RoboDK station: Robotic_Paint_Station.rdk

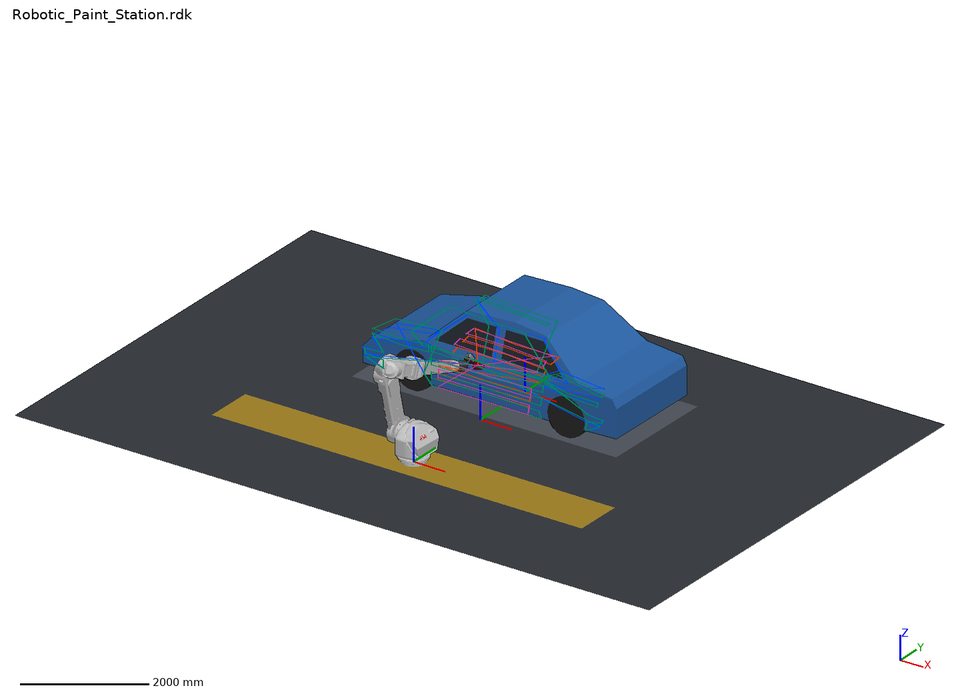
[picture v0: the station drawn from its stored meshes, robots at their saved joint values, targets as dots, program paths as lines]
Station Robotic_Paint_Station (saved by RoboDK 6.1.1). Poses are relative to the parent item; angles as X-Y-Z fixed-axis rotations.
  - frame ABB IRB 5500-27 Base at (0, 0, 0) mm
    - robot ABB IRB 5500-27: 6 axes, payload 16 kg, reach 2200 mm, repeatability 0.15 mm, weight 600 kg
        modified DH rows (alpha deg, a mm, theta deg, d mm): 0, 0, 0, 436; -90, 0, -90, -5; 0, 1300, 0, 0; -90, 0, -90, 1510.5; 35, 0, 0, 79.169; -70, 0, 180, 79.169
        base shift (0, 0, 0) mm, rotated rx 0 ry 0 rz 90 deg
        joint limits [-104, -65, -70, -719, -719, -720] to [104, 150, 70, 719, 719, 720]; home [0, 0, 0, 0, 0, 0]; saved at [-2.48, -13.69, 32.15, 0, -13.46, 0]
      - tool Generic Paint Sprayer, TCP at (50, 0, 450) mm, rotated rx 0 ry 30 rz 0 deg, size 277.6 x 203.2 x 501.7 mm
    - target Target_Home (joint target) at (1.1, 1730.94, 958.32) mm, rotated rx -169.53 ry 40.3 rz -74.78 deg; joints [-2.48, -13.69, 32.15, 0, -13.46, 0] of ABB IRB 5500-27
    - target S1_Nose1_1 (joint target) at (-2225.6, 1859.63, 480.04) mm, rotated rx -168.57 ry 36.07 rz -20.39 deg; joints [48.24, 45, -22.8, 0, -17.2, 0] of ABB IRB 5500-27
    - target S1_Nose1_2 (joint target) at (-1907.83, 1928.66, 303.01) mm, rotated rx -168.29 ry 28.55 rz -20.69 deg; joints [41.89, 41.39, -12.43, 0, -23.96, 0] of ABB IRB 5500-27
    - target S1_Nose2_1 (joint target) at (-1919.89, 1941.1, 437.66) mm, rotated rx -168.2 ry 31.78 rz -22.89 deg; joints [42.24, 38.97, -12.94, 0, -21.03, 0] of ABB IRB 5500-27
    - target S1_Nose2_2 (joint target) at (-2244.13, 1875.41, 534.28) mm, rotated rx -168.88 ry 37.79 rz -21.66 deg; joints [48.42, 45, -24.32, 0, -15.68, 0] of ABB IRB 5500-27
    - target S1_Nose3_1 (joint target) at (-2263.28, 1891.47, 594.89) mm, rotated rx -169.35 ry 39.69 rz -23.13 deg; joints [48.62, 45, -26, 0, -14, 0] of ABB IRB 5500-27
    - target S1_Nose3_2 (joint target) at (-1928.2, 1948.92, 572.22) mm, rotated rx -168.43 ry 35.06 rz -25.19 deg; joints [42.6, 36.63, -13.53, 0, -18.1, 0] of ABB IRB 5500-27
    - target S1_Fender1_1 (joint target) at (-2132.11, 1933.06, 785.84) mm, rotated rx -172.79 ry 43.01 rz -31.51 deg; joints [46.91, 38.63, -22.17, 0, -8.47, 0] of ABB IRB 5500-27
    - target S1_Fender1_2 (joint target) at (-1563.54, 1911, 817.41) mm, rotated rx -170.8 ry 37.89 rz -35.8 deg; joints [37.63, 21.02, 0.04, 0, -13.06, 0] of ABB IRB 5500-27
    - target S1_Fender1_3 (joint target) at (-1047.76, 1968.31, 876.28) mm, rotated rx -170.74 ry 37.66 rz -47.06 deg; joints [26.16, 10.19, 11.07, 0, -13.26, 0] of ABB IRB 5500-27
    - target S1_Fender2_1 (joint target) at (-1048.74, 1970.29, 928.11) mm, rotated rx -171.19 ry 39.18 rz -48.26 deg; joints [26.36, 9.37, 10.53, 0, -11.91, 0] of ABB IRB 5500-27
    - target S1_Fender2_2 (joint target) at (-1558.2, 1904.4, 868.6) mm, rotated rx -171.19 ry 39.18 rz -36.84 deg; joints [37.78, 19.8, 0.1, 0, -11.91, 0] of ABB IRB 5500-27
    - target S1_Fender2_3 (joint target) at (-2137.64, 1937.76, 836.26) mm, rotated rx -173.53 ry 44.35 rz -32.83 deg; joints [47.06, 38.23, -22.99, 0, -7.24, 0] of ABB IRB 5500-27
    - target S1_Hood1_1 (joint target) at (-1967.23, 2183.01, 902.81) mm, rotated rx 167.04 ry 45.87 rz -65.7 deg; joints [43.65, 39.99, -27.38, 0, 13.39, 0] of ABB IRB 5500-27
    - target S1_Hood1_2 (joint target) at (-1102.55, 2153.25, 1034.68) mm, rotated rx 171.5 ry 43.17 rz -74.96 deg; joints [28.61, 15.58, 0.52, 0, 9.89, 0] of ABB IRB 5500-27
    - target S1_Hood2_1 (joint target) at (-1066.31, 2257.69, 1058.44) mm, rotated rx 166.47 ry 43.43 rz -83.71 deg; joints [27.44, 18.68, -3.93, 0, 15.25, 0] of ABB IRB 5500-27
    - target S1_Hood2_2 (joint target) at (-1931.79, 2300.04, 919.17) mm, rotated rx 160.55 ry 45.99 rz -76.07 deg; joints [42.26, 43.19, -32.52, 0, 19.33, 0] of ABB IRB 5500-27
    - target S1_Ret_Door (joint target) at (-1033.89, 1758.65, 540.3) mm, rotated rx -168.52 ry 26.36 rz -34.41 deg; joints [26.42, 10.19, 20.8, 0, -26, 0] of ABB IRB 5500-27
    - target S1_Door1_1 (joint target) at (-995.1, 1908.68, 283.69) mm, rotated rx -169.9 ry 20.28 rz -33.02 deg; joints [22.91, 21.93, 14.91, 0, -31.84, 0] of ABB IRB 5500-27
    - target S1_Door1_2 (joint target) at (36.7, 1939.09, 273.54) mm, rotated rx -170.65 ry 18.19 rz -60.68 deg; joints [-6.53, 14.63, 24.32, 0, -33.95, 0] of ABB IRB 5500-27
    - target S1_Door1_3 (joint target) at (1078.9, 1931.68, 272.33) mm, rotated rx -169.79 ry 20.63 rz -89.85 deg; joints [-33.64, 24.38, 12.11, 0, -31.5, 0] of ABB IRB 5500-27
    - target S1_Door2_1 (joint target) at (1062.05, 1900.58, 393.84) mm, rotated rx -169.07 ry 23.31 rz -91.79 deg; joints [-33.37, 19.55, 14.32, 0, -28.87, 0] of ABB IRB 5500-27
    - target S1_Door2_2 (joint target) at (37.2, 1952.51, 380.39) mm, rotated rx -169.61 ry 21.25 rz -62.77 deg; joints [-6.05, 11.55, 24.33, 0, -30.89, 0] of ABB IRB 5500-27
    - target S1_Door2_3 (joint target) at (-992.52, 1905.05, 398.3) mm, rotated rx -169.11 ry 23.17 rz -35.03 deg; joints [23.27, 18.35, 15.66, 0, -29.01, 0] of ABB IRB 5500-27
    - target S1_Door3_1 (joint target) at (-1001.43, 1922.59, 504.31) mm, rotated rx -168.55 ry 26.19 rz -37.01 deg; joints [23.7, 16.15, 15, 0, -26.15, 0] of ABB IRB 5500-27
    - target S1_Door3_2 (joint target) at (37.06, 1959.18, 488.1) mm, rotated rx -168.84 ry 24.42 rz -64.87 deg; joints [-5.56, 8.46, 24.35, 0, -27.81, 0] of ABB IRB 5500-27
    - target S1_Door3_3 (joint target) at (1072.37, 1918.91, 500.61) mm, rotated rx -168.52 ry 26.34 rz -93.77 deg; joints [-32.94, 17.41, 13.6, 0, -26.01, 0] of ABB IRB 5500-27
    - target S1_Door4_1 (joint target) at (1080.95, 1933.7, 608.41) mm, rotated rx -168.24 ry 29.44 rz -95.8 deg; joints [-32.52, 15.36, 12.79, 0, -23.15, 0] of ABB IRB 5500-27
    - target S1_Door4_2 (joint target) at (36.59, 1958.97, 596.14) mm, rotated rx -168.36 ry 27.7 rz -66.98 deg; joints [-5.07, 5.36, 24.38, 0, -24.74, 0] of ABB IRB 5500-27
    - target S1_Door4_3 (joint target) at (-1008.33, 1936.75, 611.3) mm, rotated rx -168.24 ry 29.28 rz -39.03 deg; joints [24.12, 14.04, 14.25, 0, -23.29, 0] of ABB IRB 5500-27
    - target S1_Door5_1 (joint target) at (-1014.28, 1947.2, 719.07) mm, rotated rx -168.22 ry 32.45 rz -41.11 deg; joints [24.56, 12.03, 13.4, 0, -20.43, 0] of ABB IRB 5500-27
    - target S1_Door5_2 (joint target) at (36.4, 1952.31, 704.35) mm, rotated rx -168.2 ry 31.08 rz -69.17 deg; joints [-4.59, 2.26, 24.4, 0, -21.66, 0] of ABB IRB 5500-27
    - target S1_Door5_3 (joint target) at (1087.47, 1945.07, 717.07) mm, rotated rx -168.23 ry 32.6 rz -97.89 deg; joints [-32.1, 13.4, 11.89, 0, -20.29, 0] of ABB IRB 5500-27
    - target S1_Door6_1 (joint target) at (1091.81, 1953.69, 825.52) mm, rotated rx -168.53 ry 35.79 rz -100.06 deg; joints [-31.67, 11.57, 10.88, 0, -17.45, 0] of ABB IRB 5500-27
    - target S1_Door6_2 (joint target) at (35.83, 1938.56, 811.93) mm, rotated rx -168.37 ry 34.52 rz -71.44 deg; joints [-4.1, -0.86, 24.44, 0, -18.58, 0] of ABB IRB 5500-27
    - target S1_Door6_3 (joint target) at (-1018.43, 1954.84, 827.37) mm, rotated rx -168.5 ry 35.65 rz -43.28 deg; joints [24.99, 10.14, 12.43, 0, -17.58, 0] of ABB IRB 5500-27
    - target S1_Door7_1 (joint target) at (-1021.03, 1959.35, 934.99) mm, rotated rx -169.13 ry 38.85 rz -45.59 deg; joints [25.42, 8.38, 11.36, 0, -14.74, 0] of ABB IRB 5500-27
    - target S1_Door7_2 (joint target) at (35.73, 1918.46, 918.39) mm, rotated rx -168.93 ry 37.99 rz -73.88 deg; joints [-3.62, -3.97, 24.47, 0, -15.5, 0] of ABB IRB 5500-27
    - target S1_Door7_3 (joint target) at (1094.67, 1958.91, 934.44) mm, rotated rx -169.17 ry 39 rz -102.39 deg; joints [-31.25, 9.84, 9.77, 0, -14.61, 0] of ABB IRB 5500-27
    - target S1_Ret_Pillar (joint target) at (-1047.69, 1750.88, 1005.83) mm, rotated rx -173.43 ry 41.27 rz -49.35 deg; joints [29.67, -0.19, 18.45, 0, -8.26, 0] of ABB IRB 5500-27
    - target S1_APil_1 (joint target) at (-1085.22, 2017.79, 1022.51) mm, rotated rx 176.04 ry 42.59 rz -67.35 deg; joints [29.1, 10.29, 6.96, 0, 4.76, 0] of ABB IRB 5500-27
    - target S1_APil_2 (joint target) at (-461.04, 2108.16, 1553.88) mm, rotated rx 155.15 ry 52.69 rz -106.77 deg; joints [15.38, 0, 3.11, 0, 18.89, 0] of ABB IRB 5500-27
    - target S1_Cant_1 (joint target) at (-406.96, 2128.53, 1584.57) mm, rotated rx 146.8 ry 50.14 rz -118.16 deg; joints [14.89, 0.58, 1.37, 0, 26.05, 0] of ABB IRB 5500-27
    - target S1_Cant_2 (joint target) at (334.35, 2079.2, 1576.67) mm, rotated rx 147.19 ry 50.1 rz -137.61 deg; joints [-4.98, -2.11, 4.26, 0, 25.85, 0] of ABB IRB 5500-27
    - target S1_Cant_3 (joint target) at (1068.74, 2057.28, 1601.52) mm, rotated rx 145.27 ry 50.27 rz -158.23 deg; joints [-23.55, 7.24, -6.06, 0, 26.82, 0] of ABB IRB 5500-27
    - target S1_CPil_1 (joint target) at (1034.33, 2039.03, 1569.29) mm, rotated rx 153.95 ry 52.94 rz -147.41 deg; joints [-23.94, 5.62, -3.11, 0, 19.49, 0] of ABB IRB 5500-27
    - target S1_CPil_2 (joint target) at (1621.44, 1846.13, 1053.12) mm, rotated rx 174.14 ry 44.25 rz -139.45 deg; joints [-40.27, 16.89, -1.48, 0, 6.59, 0] of ABB IRB 5500-27
    - target S1_Ret_BPil (joint target) at (549.31, 1741.35, 1184.47) mm, rotated rx -177.48 ry 47.41 rz -104.09 deg; joints [-17.82, -12.59, 25.12, 0, -2.53, 0] of ABB IRB 5500-27
    - target S1_BPil_1 (joint target) at (186.88, 1914.62, 996.74) mm, rotated rx -178.08 ry 41.55 rz -92.64 deg; joints [-5.85, -5.35, 23.76, 0, -2.41, 0] of ABB IRB 5500-27
    - target S1_BPil_2 (joint target) at (186.93, 2066.73, 1500.15) mm, rotated rx 165.22 ry 53.82 rz -112.49 deg; joints [-3.2, -3.64, 8.35, 0, 11.29, 0] of ABB IRB 5500-27
    - target S1_Roof1_1 (joint target) at (-460.71, 2348.38, 1749.55) mm, rotated rx 122.28 ry 33.89 rz -147.32 deg; joints [17.76, 12.35, -17.99, 0, 53.63, 0] of ABB IRB 5500-27
    - target S1_Roof1_2 (joint target) at (964.63, 2213.74, 1745.81) mm, rotated rx 122.22 ry 33.86 rz 177.92 deg; joints [-16.94, 13.34, -19.02, 0, 53.68, 0] of ABB IRB 5500-27
    - target S1_Roof2_1 (joint target) at (967.48, 2302.77, 1719.45) mm, rotated rx 120.57 ry 30.14 rz 175.73 deg; joints [-16.06, 17.59, -23.78, 0, 58.19, 0] of ABB IRB 5500-27
    - target S1_Roof2_2 (joint target) at (-436.75, 2431.34, 1724.45) mm, rotated rx 120.72 ry 30.21 rz -151.1 deg; joints [16.98, 16.3, -22.38, 0, 58.08, 0] of ABB IRB 5500-27
    - target S1_Roof3_1 (joint target) at (-442.87, 2593.03, 1710.21) mm, rotated rx 117.22 ry 25.16 rz -156.15 deg; joints [16.46, 24.63, -32.92, 0, 64.29, 0] of ABB IRB 5500-27
    - target S1_Roof3_2 (joint target) at (986.3, 2476.69, 1712.68) mm, rotated rx 116.42 ry 24.66 rz 171.76 deg; joints [-15, 26.49, -35.44, 0, 64.95, 0] of ABB IRB 5500-27
    - target S1_Ret_Rear (joint target) at (1089.9, 1709.82, 1074.98) mm, rotated rx -174.56 ry 43.36 rz -114.73 deg; joints [-33.43, -1.82, 18.16, 0, -6.34, 0] of ABB IRB 5500-27
    - target S1_Trnk1_1 (joint target) at (1286.21, 2128.18, 1086.31) mm, rotated rx 167.41 ry 44.29 rz -138.57 deg; joints [-29.17, 17.87, -3.69, 0, 13.81, 0] of ABB IRB 5500-27
    - target S1_Trnk1_2 (joint target) at (2138.82, 2113.18, 1005.84) mm, rotated rx 159.08 ry 47.76 rz -162.55 deg; joints [-43.11, 42.46, -33.83, 0, 19.37, 0] of ABB IRB 5500-27
    - target S1_Qtr1_1 (joint target) at (1108.2, 1947.47, 813.97) mm, rotated rx -170.31 ry 35.92 rz -103.38 deg; joints [-31.73, 11.81, 11.01, 0, -14.83, 0] of ABB IRB 5500-27
    - target S1_Qtr1_2 (joint target) at (1605.25, 1889.84, 818.76) mm, rotated rx -170.84 ry 38.03 rz -115.54 deg; joints [-41.98, 21.42, -0.49, 0, -12.93, 0] of ABB IRB 5500-27
    - target S1_Qtr1_3 (joint target) at (2162.61, 1911.94, 846.58) mm, rotated rx -173.68 ry 44.62 rz -129.42 deg; joints [-49.24, 38.15, -23.16, 0, -7, 0] of ABB IRB 5500-27
    - target S1_Qtr2_1 (joint target) at (2169.44, 1917.68, 917.73) mm, rotated rx -174.91 ry 46.51 rz -131.41 deg; joints [-49.04, 37.63, -24.37, 0, -5.26, 0] of ABB IRB 5500-27
    - target S1_Qtr2_2 (joint target) at (1598.86, 1881.54, 911.67) mm, rotated rx -171.65 ry 40.43 rz -117.54 deg; joints [-41.71, 19.45, -0.67, 0, -10.78, 0] of ABB IRB 5500-27
    - target S1_Qtr2_3 (joint target) at (1110.87, 1952.75, 927.55) mm, rotated rx -171.22 ry 39.24 rz -105.96 deg; joints [-31.28, 9.99, 9.86, 0, -11.85, 0] of ABB IRB 5500-27
    - target S1_RSk1_1 (joint target) at (1928.28, 1948.84, 572.22) mm, rotated rx -168.43 ry 35.06 rz -114.58 deg; joints [-46.79, 36.63, -13.53, 0, -18.1, 0] of ABB IRB 5500-27
    - target S1_RSk1_2 (joint target) at (2237.47, 1894.83, 577.43) mm, rotated rx -169.14 ry 38.91 rz -122.38 deg; joints [-51.32, 44.53, -24.84, 0, -14.69, 0] of ABB IRB 5500-27
    - target S1_RSk2_1 (joint target) at (2218.08, 1878.01, 493.19) mm, rotated rx -168.64 ry 36.49 rz -120.56 deg; joints [-51.58, 45, -23.17, 0, -16.83, 0] of ABB IRB 5500-27
    - target S1_RSk2_2 (joint target) at (1920.22, 1940.78, 437.66) mm, rotated rx -168.2 ry 31.78 rz -112.27 deg; joints [-47.14, 38.97, -12.94, 0, -21.03, 0] of ABB IRB 5500-27
    - target S1_RSk3_1 (joint target) at (1907.9, 1928.59, 303.01) mm, rotated rx -168.29 ry 28.55 rz -110.07 deg; joints [-47.49, 41.39, -12.43, 0, -23.96, 0] of ABB IRB 5500-27
    - target S1_RSk3_2 (joint target) at (2200.11, 1863.41, 444.32) mm, rotated rx -168.42 ry 34.93 rz -119.42 deg; joints [-51.74, 45, -21.79, 0, -18.21, 0] of ABB IRB 5500-27
    - target S2_Bmp1_1 (joint target) at (-855.22, 1891.67, 297.5) mm, rotated rx -170.03 ry 19.91 rz -36.14 deg; joints [19.48, 18.78, 18.43, 0, -32.21, 0] of ABB IRB 5500-27
    - target S2_Bmp1_2 (joint target) at (0.46, 1939.19, 273.26) mm, rotated rx -170.65 ry 18.19 rz -59.62 deg; joints [-5.46, 14.63, 24.33, 0, -33.95, 0] of ABB IRB 5500-27
    - target S2_Bmp1_3 (joint target) at (855.37, 1891.6, 297.5) mm, rotated rx -170.03 ry 19.91 rz -84.8 deg; joints [-29.18, 18.78, 18.43, 0, -32.21, 0] of ABB IRB 5500-27
    - target S2_Bmp2_1 (joint target) at (863.55, 1908.53, 410.17) mm, rotated rx -169.14 ry 23.04 rz -86.92 deg; joints [-28.72, 16.02, 18.11, 0, -29.13, 0] of ABB IRB 5500-27
    - target S2_Bmp2_2 (joint target) at (0.82, 1952.91, 385.38) mm, rotated rx -169.57 ry 21.39 rz -61.81 deg; joints [-4.96, 11.39, 24.35, 0, -30.74, 0] of ABB IRB 5500-27
    - target S2_Bmp2_3 (joint target) at (-862.53, 1908.99, 410.17) mm, rotated rx -169.14 ry 23.04 rz -38.26 deg; joints [19.94, 16.02, 18.11, 0, -29.13, 0] of ABB IRB 5500-27
    - target S2_Bmp3_1 (joint target) at (-868.79, 1923.35, 521.8) mm, rotated rx -168.54 ry 26.25 rz -40.36 deg; joints [20.4, 13.47, 17.62, 0, -26.09, 0] of ABB IRB 5500-27
    - target S2_Bmp3_2 (joint target) at (0.61, 1959.4, 498.36) mm, rotated rx -168.78 ry 24.73 rz -64 deg; joints [-4.45, 8.15, 24.37, 0, -27.52, 0] of ABB IRB 5500-27
    - target S2_Bmp3_3 (joint target) at (870.2, 1922.71, 521.8) mm, rotated rx -168.54 ry 26.25 rz -89.02 deg; joints [-28.26, 13.47, 17.62, 0, -26.09, 0] of ABB IRB 5500-27
    - target S2_Bmp4_1 (joint target) at (875.37, 1934.23, 632.46) mm, rotated rx -168.23 ry 29.5 rz -91.13 deg; joints [-27.8, 11.12, 16.97, 0, -23.09, 0] of ABB IRB 5500-27
    - target S2_Bmp4_2 (joint target) at (0.27, 1958.61, 611.63) mm, rotated rx -168.32 ry 28.18 rz -66.22 deg; joints [-3.94, 4.91, 24.39, 0, -24.3, 0] of ABB IRB 5500-27
    - target S2_Bmp4_3 (joint target) at (-874.02, 1934.84, 632.46) mm, rotated rx -168.23 ry 29.5 rz -42.47 deg; joints [20.86, 11.12, 16.97, 0, -23.09, 0] of ABB IRB 5500-27
    - target S2_Bonnet1_1 (joint target) at (917.87, 2057.79, 801.97) mm, rotated rx -177.87 ry 36.68 rz -110.36 deg; joints [-24.4, 12.34, 10.92, 0, -3.25, 0] of ABB IRB 5500-27
    - target S2_Bonnet1_2 (joint target) at (87.25, 2076.19, 805.31) mm, rotated rx -177.52 ry 36.03 rz -88.12 deg; joints [-2.9, 4.98, 18.91, 0, -3.88, 0] of ABB IRB 5500-27
    - target S2_Bonnet1_3 (joint target) at (-754.4, 2123.18, 801.97) mm, rotated rx -177.87 ry 36.68 rz -66.76 deg; joints [19.2, 12.34, 10.92, 0, -3.25, 0] of ABB IRB 5500-27
    - target S2_Bonnet2_1 (joint target) at (-725.24, 2238.59, 874.14) mm, rotated rx 177.64 ry 39.18 rz -75.64 deg; joints [18.54, 15.16, 5.59, 0, 3.25, 0] of ABB IRB 5500-27
    - target S2_Bonnet2_2 (joint target) at (111.75, 2222.36, 878.86) mm, rotated rx 178.14 ry 38.59 rz -95.7 deg; joints [-2.35, 9.78, 11.59, 0, 2.63, 0] of ABB IRB 5500-27
    - target S2_Bonnet2_3 (joint target) at (934.51, 2159.62, 874.14) mm, rotated rx 177.64 ry 39.18 rz -116.99 deg; joints [-22.81, 15.16, 5.59, 0, 3.25, 0] of ABB IRB 5500-27
    - target S2_Bonnet3_1 (joint target) at (944.55, 2242.71, 946.45) mm, rotated rx 172.26 ry 41.11 rz -124.32 deg; joints [-21.37, 17.42, 0.81, 0, 9.76, 0] of ABB IRB 5500-27
    - target S2_Bonnet3_2 (joint target) at (135.36, 2332.26, 948.62) mm, rotated rx 172.92 ry 40.57 rz -103.9 deg; joints [-1.88, 13.33, 5.54, 0, 9.14, 0] of ABB IRB 5500-27
    - target S2_Bonnet3_3 (joint target) at (-689.97, 2333.64, 946.45) mm, rotated rx 172.26 ry 41.11 rz -85.01 deg; joints [17.94, 17.42, 0.81, 0, 9.76, 0] of ABB IRB 5500-27
    - target S2_Bonnet4_1 (joint target) at (-662.58, 2445.82, 1008.58) mm, rotated rx 165.99 ry 42.36 rz -94.91 deg; joints [17.43, 20.92, -5.3, 0, 16.38, 0] of ABB IRB 5500-27
    - target S2_Bonnet4_2 (joint target) at (158.03, 2415.68, 1019.07) mm, rotated rx 166.9 ry 41.86 rz -112.64 deg; joints [-1.46, 16, 0.33, 0, 15.67, 0] of ABB IRB 5500-27
    - target S2_Bonnet4_3 (joint target) at (961.21, 2344.59, 1008.58) mm, rotated rx 165.99 ry 42.36 rz -132.36 deg; joints [-20.02, 20.92, -5.3, 0, 16.38, 0] of ABB IRB 5500-27
    - target S2_Bonnet5_1 (joint target) at (993, 2515.38, 1064.78) mm, rotated rx 158.52 ry 43.53 rz -141.02 deg; joints [-18.64, 27.82, -15.76, 0, 22.94, 0] of ABB IRB 5500-27
    - target S2_Bonnet5_2 (joint target) at (174.44, 2508.6, 1063.51) mm, rotated rx 161.75 ry 42.39 rz -119.67 deg; joints [-1.13, 19.56, -5.31, 0, 20.75, 0] of ABB IRB 5500-27
    - target S2_Bonnet5_3 (joint target) at (-664.17, 2621.46, 1064.78) mm, rotated rx 158.52 ry 43.53 rz -105.26 deg; joints [17.12, 27.82, -15.76, 0, 22.94, 0] of ABB IRB 5500-27
    - target S3_RSk1_1 (joint target) at (-2200.33, 1863.16, 444.32) mm, rotated rx -168.42 ry 34.93 rz -19.94 deg; joints [47.74, 45, -21.79, 0, -18.21, 0] of ABB IRB 5500-27
    - target S3_RSk1_2 (joint target) at (-1907.83, 1928.66, 303.01) mm, rotated rx -168.29 ry 28.55 rz -20.69 deg; joints [41.89, 41.39, -12.43, 0, -23.96, 0] of ABB IRB 5500-27
    - target S3_RSk2_1 (joint target) at (-1919.89, 1941.1, 437.66) mm, rotated rx -168.2 ry 31.78 rz -22.89 deg; joints [42.24, 38.97, -12.94, 0, -21.03, 0] of ABB IRB 5500-27
    - target S3_RSk2_2 (joint target) at (-2218.02, 1878.09, 493.19) mm, rotated rx -168.64 ry 36.49 rz -21.07 deg; joints [47.91, 45, -23.17, 0, -16.83, 0] of ABB IRB 5500-27
    - target S3_RSk3_1 (joint target) at (-2237.47, 1894.83, 577.43) mm, rotated rx -169.14 ry 38.91 rz -22.9 deg; joints [48.16, 44.53, -24.84, 0, -14.69, 0] of ABB IRB 5500-27
    - target S3_RSk3_2 (joint target) at (-1928.2, 1948.92, 572.22) mm, rotated rx -168.43 ry 35.06 rz -25.19 deg; joints [42.6, 36.63, -13.53, 0, -18.1, 0] of ABB IRB 5500-27
    - target S3_Qtr1_1 (joint target) at (-2138.72, 1938.62, 846.58) mm, rotated rx -173.68 ry 44.62 rz -33.09 deg; joints [47.09, 38.15, -23.16, 0, -7, 0] of ABB IRB 5500-27
    - target S3_Qtr1_2 (joint target) at (-1579.38, 1911.52, 818.76) mm, rotated rx -170.84 ry 38.03 rz -35.63 deg; joints [37.93, 21.42, -0.49, 0, -12.93, 0] of ABB IRB 5500-27
    - target S3_Qtr1_3 (joint target) at (-1077.01, 1964.9, 813.97) mm, rotated rx -170.31 ry 35.92 rz -45.01 deg; joints [26.64, 11.81, 11.01, 0, -14.83, 0] of ABB IRB 5500-27
    - target S3_Qtr2_1 (joint target) at (-1079.76, 1970.13, 927.55) mm, rotated rx -171.22 ry 39.24 rz -47.6 deg; joints [27.08, 9.99, 9.86, 0, -11.85, 0] of ABB IRB 5500-27
    - target S3_Qtr2_2 (joint target) at (-1572.32, 1903.77, 911.67) mm, rotated rx -171.65 ry 40.43 rz -37.63 deg; joints [38.2, 19.45, -0.67, 0, -10.78, 0] of ABB IRB 5500-27
    - target S3_Qtr2_3 (joint target) at (-2145.18, 1944.78, 917.73) mm, rotated rx -174.91 ry 46.51 rz -35.08 deg; joints [47.29, 37.63, -24.37, 0, -5.26, 0] of ABB IRB 5500-27
    - target S3_Trnk1_1 (joint target) at (-1942.46, 2294.97, 1005.84) mm, rotated rx 159.08 ry 47.76 rz -76.96 deg; joints [42.48, 42.46, -33.83, 0, 19.37, 0] of ABB IRB 5500-27
    - target S3_Trnk1_2 (joint target) at (-1047.47, 2255.28, 1086.31) mm, rotated rx 167.41 ry 44.29 rz -82.51 deg; joints [26.89, 17.87, -3.69, 0, 13.81, 0] of ABB IRB 5500-27
    - target S3_Ret_Door (joint target) at (-1033.89, 1758.65, 540.3) mm, rotated rx -168.52 ry 26.36 rz -34.41 deg; joints [26.42, 10.19, 20.8, 0, -26, 0] of ABB IRB 5500-27
    - target S3_Door1_1 (joint target) at (-995.1, 1908.68, 283.69) mm, rotated rx -169.9 ry 20.28 rz -33.02 deg; joints [22.91, 21.93, 14.91, 0, -31.84, 0] of ABB IRB 5500-27
    - target S3_Door1_2 (joint target) at (36.7, 1939.09, 273.54) mm, rotated rx -170.65 ry 18.19 rz -60.68 deg; joints [-6.53, 14.63, 24.32, 0, -33.95, 0] of ABB IRB 5500-27
    - target S3_Door1_3 (joint target) at (1078.9, 1931.68, 272.33) mm, rotated rx -169.79 ry 20.63 rz -89.85 deg; joints [-33.64, 24.38, 12.11, 0, -31.5, 0] of ABB IRB 5500-27
    - target S3_Door2_1 (joint target) at (1062.05, 1900.58, 393.84) mm, rotated rx -169.07 ry 23.31 rz -91.79 deg; joints [-33.37, 19.55, 14.32, 0, -28.87, 0] of ABB IRB 5500-27
    - target S3_Door2_2 (joint target) at (37.2, 1952.51, 380.39) mm, rotated rx -169.61 ry 21.25 rz -62.77 deg; joints [-6.05, 11.55, 24.33, 0, -30.89, 0] of ABB IRB 5500-27
    - target S3_Door2_3 (joint target) at (-992.52, 1905.05, 398.3) mm, rotated rx -169.11 ry 23.17 rz -35.03 deg; joints [23.27, 18.35, 15.66, 0, -29.01, 0] of ABB IRB 5500-27
    - target S3_Door3_1 (joint target) at (-1001.43, 1922.59, 504.31) mm, rotated rx -168.55 ry 26.19 rz -37.01 deg; joints [23.7, 16.15, 15, 0, -26.15, 0] of ABB IRB 5500-27
    - target S3_Door3_2 (joint target) at (37.06, 1959.18, 488.1) mm, rotated rx -168.84 ry 24.42 rz -64.87 deg; joints [-5.56, 8.46, 24.35, 0, -27.81, 0] of ABB IRB 5500-27
    - target S3_Door3_3 (joint target) at (1072.37, 1918.91, 500.61) mm, rotated rx -168.52 ry 26.34 rz -93.77 deg; joints [-32.94, 17.41, 13.6, 0, -26.01, 0] of ABB IRB 5500-27
    - target S3_Door4_1 (joint target) at (1080.95, 1933.7, 608.41) mm, rotated rx -168.24 ry 29.44 rz -95.8 deg; joints [-32.52, 15.36, 12.79, 0, -23.15, 0] of ABB IRB 5500-27
    - target S3_Door4_2 (joint target) at (36.59, 1958.97, 596.14) mm, rotated rx -168.36 ry 27.7 rz -66.98 deg; joints [-5.07, 5.36, 24.38, 0, -24.74, 0] of ABB IRB 5500-27
    - target S3_Door4_3 (joint target) at (-1008.33, 1936.75, 611.3) mm, rotated rx -168.24 ry 29.28 rz -39.03 deg; joints [24.12, 14.04, 14.25, 0, -23.29, 0] of ABB IRB 5500-27
    - target S3_Door5_1 (joint target) at (-1014.28, 1947.2, 719.07) mm, rotated rx -168.22 ry 32.45 rz -41.11 deg; joints [24.56, 12.03, 13.4, 0, -20.43, 0] of ABB IRB 5500-27
    - target S3_Door5_2 (joint target) at (36.4, 1952.31, 704.35) mm, rotated rx -168.2 ry 31.08 rz -69.17 deg; joints [-4.59, 2.26, 24.4, 0, -21.66, 0] of ABB IRB 5500-27
    - target S3_Door5_3 (joint target) at (1087.47, 1945.07, 717.07) mm, rotated rx -168.23 ry 32.6 rz -97.89 deg; joints [-32.1, 13.4, 11.89, 0, -20.29, 0] of ABB IRB 5500-27
    - target S3_Door6_1 (joint target) at (1091.81, 1953.69, 825.52) mm, rotated rx -168.53 ry 35.79 rz -100.06 deg; joints [-31.67, 11.57, 10.88, 0, -17.45, 0] of ABB IRB 5500-27
    - target S3_Door6_2 (joint target) at (35.83, 1938.56, 811.93) mm, rotated rx -168.37 ry 34.52 rz -71.44 deg; joints [-4.1, -0.86, 24.44, 0, -18.58, 0] of ABB IRB 5500-27
    - target S3_Door6_3 (joint target) at (-1018.43, 1954.84, 827.37) mm, rotated rx -168.5 ry 35.65 rz -43.28 deg; joints [24.99, 10.14, 12.43, 0, -17.58, 0] of ABB IRB 5500-27
    - target S3_Door7_1 (joint target) at (-1021.03, 1959.35, 934.99) mm, rotated rx -169.13 ry 38.85 rz -45.59 deg; joints [25.42, 8.38, 11.36, 0, -14.74, 0] of ABB IRB 5500-27
    - target S3_Door7_2 (joint target) at (35.73, 1918.46, 918.39) mm, rotated rx -168.93 ry 37.99 rz -73.88 deg; joints [-3.62, -3.97, 24.47, 0, -15.5, 0] of ABB IRB 5500-27
    - target S3_Door7_3 (joint target) at (1094.67, 1958.91, 934.44) mm, rotated rx -169.17 ry 39 rz -102.39 deg; joints [-31.25, 9.84, 9.77, 0, -14.61, 0] of ABB IRB 5500-27
    - target S3_Ret_Pillar (joint target) at (-1047.69, 1750.88, 1005.83) mm, rotated rx -173.43 ry 41.27 rz -49.35 deg; joints [29.67, -0.19, 18.45, 0, -8.26, 0] of ABB IRB 5500-27
    - target S3_CPil_1 (joint target) at (-1430.22, 1978.96, 1053.01) mm, rotated rx 174.26 ry 44.15 rz -62.14 deg; joints [36.87, 16.24, -0.71, 0, 6.48, 0] of ABB IRB 5500-27
    - target S3_CPil_2 (joint target) at (-832.81, 2115.56, 1567.58) mm, rotated rx 154.11 ry 52.91 rz -98.85 deg; joints [24.45, 5.06, -2.47, 0, 19.41, 0] of ABB IRB 5500-27
    - target S3_Cant_1 (joint target) at (-786.79, 2158.6, 1600.07) mm, rotated rx 145.48 ry 50.25 rz -110.51 deg; joints [23.95, 6.32, -5.03, 0, 26.72, 0] of ABB IRB 5500-27
    - target S3_Cant_2 (joint target) at (-44, 2102.04, 1576.18) mm, rotated rx 147.21 ry 50.1 rz -127.24 deg; joints [5.36, -2.26, 4.42, 0, 25.84, 0] of ABB IRB 5500-27
    - target S3_Cant_3 (joint target) at (679.07, 2063.2, 1584.86) mm, rotated rx 146.78 ry 50.14 rz -147.23 deg; joints [-14.16, 0.8, 1.14, 0, 26.06, 0] of ABB IRB 5500-27
    - target S3_APil_1 (joint target) at (670.38, 2057.22, 1554.59) mm, rotated rx 155.11 ry 52.7 rz -137.2 deg; joints [-15.01, 0.25, 2.84, 0, 18.91, 0] of ABB IRB 5500-27
    - target S3_APil_2 (joint target) at (1237.64, 1917.14, 1022.63) mm, rotated rx 176.08 ry 42.55 rz -128.41 deg; joints [-32.02, 9.9, 7.39, 0, 4.72, 0] of ABB IRB 5500-27
    - target S3_Ret_BPil (joint target) at (446.76, 1748.11, 1185.35) mm, rotated rx -177.63 ry 47.59 rz -101.13 deg; joints [-14.62, -13.64, 26, 0, -2.36, 0] of ABB IRB 5500-27
    - target S3_BPil_1 (joint target) at (-17.23, 1922.19, 996.95) mm, rotated rx -178.09 ry 41.56 rz -86.56 deg; joints [0.24, -5.42, 23.82, 0, -2.4, 0] of ABB IRB 5500-27
    - target S3_BPil_2 (joint target) at (-17.37, 2071.93, 1499.95) mm, rotated rx 165.23 ry 53.83 rz -106.83 deg; joints [2.45, -3.78, 8.49, 0, 11.28, 0] of ABB IRB 5500-27
    - target S3_Roof1_1 (joint target) at (-460.71, 2348.38, 1749.55) mm, rotated rx 122.28 ry 33.89 rz -147.32 deg; joints [17.76, 12.35, -17.99, 0, 53.63, 0] of ABB IRB 5500-27
    - target S3_Roof1_2 (joint target) at (964.63, 2213.74, 1745.81) mm, rotated rx 122.22 ry 33.86 rz 177.92 deg; joints [-16.94, 13.34, -19.02, 0, 53.68, 0] of ABB IRB 5500-27
    - target S3_Roof2_1 (joint target) at (967.48, 2302.77, 1719.45) mm, rotated rx 120.57 ry 30.14 rz 175.73 deg; joints [-16.06, 17.59, -23.78, 0, 58.19, 0] of ABB IRB 5500-27
    - target S3_Roof2_2 (joint target) at (-436.75, 2431.34, 1724.45) mm, rotated rx 120.72 ry 30.21 rz -151.1 deg; joints [16.98, 16.3, -22.38, 0, 58.08, 0] of ABB IRB 5500-27
    - target S3_Roof3_1 (joint target) at (-442.87, 2593.03, 1710.21) mm, rotated rx 117.22 ry 25.16 rz -156.15 deg; joints [16.46, 24.63, -32.92, 0, 64.29, 0] of ABB IRB 5500-27
    - target S3_Roof3_2 (joint target) at (986.3, 2476.69, 1712.68) mm, rotated rx 116.42 ry 24.66 rz 171.76 deg; joints [-15, 26.49, -35.44, 0, 64.95, 0] of ABB IRB 5500-27
    - target S3_Ret_Front (joint target) at (1089.9, 1709.82, 1074.98) mm, rotated rx -174.56 ry 43.36 rz -114.73 deg; joints [-33.43, -1.82, 18.16, 0, -6.34, 0] of ABB IRB 5500-27
    - target S3_Hood1_1 (joint target) at (1323.43, 2117.24, 1058.44) mm, rotated rx 166.47 ry 43.43 rz -141 deg; joints [-29.85, 18.68, -3.93, 0, 15.25, 0] of ABB IRB 5500-27
    - target S3_Hood1_2 (joint target) at (2145.06, 2102.55, 919.17) mm, rotated rx 160.55 ry 45.99 rz -161.67 deg; joints [-43.34, 43.19, -32.52, 0, 19.33, 0] of ABB IRB 5500-27
    - target S3_Hood2_1 (joint target) at (2143.79, 2009.9, 902.81) mm, rotated rx 167.04 ry 45.87 rz -154.57 deg; joints [-45.22, 39.99, -27.38, 0, 13.39, 0] of ABB IRB 5500-27
    - target S3_Hood2_2 (joint target) at (1316.68, 2029.4, 1034.68) mm, rotated rx 171.5 ry 43.17 rz -135.05 deg; joints [-31.48, 15.58, 0.52, 0, 9.89, 0] of ABB IRB 5500-27
    - target S3_Fend1_1 (joint target) at (1110.19, 1950.79, 875.85) mm, rotated rx -170.76 ry 37.73 rz -104.77 deg; joints [-31.49, 10.81, 10.39, 0, -13.2, 0] of ABB IRB 5500-27
    - target S3_Fend1_2 (joint target) at (1605.25, 1889.84, 818.76) mm, rotated rx -170.84 ry 38.03 rz -115.54 deg; joints [-41.98, 21.42, -0.49, 0, -12.93, 0] of ABB IRB 5500-27
    - target S3_Fend1_3 (joint target) at (2156.02, 1906.36, 785.84) mm, rotated rx -172.79 ry 43.01 rz -127.83 deg; joints [-49.41, 38.63, -22.17, 0, -8.47, 0] of ABB IRB 5500-27
    - target S3_Fend2_1 (joint target) at (2161.63, 1910.96, 836.26) mm, rotated rx -173.53 ry 44.35 rz -129.16 deg; joints [-49.27, 38.23, -22.99, 0, -7.24, 0] of ABB IRB 5500-27
    - target S3_Fend2_2 (joint target) at (1597.41, 1880.17, 868.32) mm, rotated rx -171.22 ry 39.24 rz -116.53 deg; joints [-41.85, 20.07, -0.22, 0, -11.85, 0] of ABB IRB 5500-27
    - target S3_Fend2_3 (joint target) at (1110.87, 1952.75, 927.55) mm, rotated rx -171.22 ry 39.24 rz -105.96 deg; joints [-31.28, 9.99, 9.86, 0, -11.85, 0] of ABB IRB 5500-27
    - target S3_Nose1_1 (joint target) at (1928.28, 1948.84, 572.22) mm, rotated rx -168.43 ry 35.06 rz -114.58 deg; joints [-46.79, 36.63, -13.53, 0, -18.1, 0] of ABB IRB 5500-27
    - target S3_Nose1_2 (joint target) at (2263.35, 1891.38, 594.89) mm, rotated rx -169.35 ry 39.69 rz -123.36 deg; joints [-51.61, 45, -26, 0, -14, 0] of ABB IRB 5500-27
    - target S3_Nose2_1 (joint target) at (2244.16, 1875.39, 534.28) mm, rotated rx -168.88 ry 37.79 rz -121.89 deg; joints [-51.81, 45, -24.32, 0, -15.68, 0] of ABB IRB 5500-27
    - target S3_Nose2_2 (joint target) at (1920.22, 1940.78, 437.66) mm, rotated rx -168.2 ry 31.78 rz -112.27 deg; joints [-47.14, 38.97, -12.94, 0, -21.03, 0] of ABB IRB 5500-27
    - target S3_Nose3_1 (joint target) at (1907.9, 1928.59, 303.01) mm, rotated rx -168.29 ry 28.55 rz -110.07 deg; joints [-47.49, 41.39, -12.43, 0, -23.96, 0] of ABB IRB 5500-27
    - target S3_Nose3_2 (joint target) at (2225.66, 1859.56, 480.04) mm, rotated rx -168.57 ry 36.07 rz -120.63 deg; joints [-52, 45, -22.8, 0, -17.2, 0] of ABB IRB 5500-27
    - target S4_RBmp1_1 (joint target) at (-855.22, 1891.67, 297.5) mm, rotated rx -170.03 ry 19.91 rz -36.14 deg; joints [19.48, 18.78, 18.43, 0, -32.21, 0] of ABB IRB 5500-27
    - target S4_RBmp1_2 (joint target) at (0.46, 1939.19, 273.26) mm, rotated rx -170.65 ry 18.19 rz -59.62 deg; joints [-5.46, 14.63, 24.33, 0, -33.95, 0] of ABB IRB 5500-27
    - target S4_RBmp1_3 (joint target) at (855.37, 1891.6, 297.5) mm, rotated rx -170.03 ry 19.91 rz -84.8 deg; joints [-29.18, 18.78, 18.43, 0, -32.21, 0] of ABB IRB 5500-27
    - target S4_RBmp2_1 (joint target) at (865.45, 1912.06, 441.14) mm, rotated rx -168.94 ry 23.92 rz -87.5 deg; joints [-28.6, 15.27, 18.02, 0, -28.29, 0] of ABB IRB 5500-27
    - target S4_RBmp2_2 (joint target) at (0.77, 1955.53, 416.17) mm, rotated rx -169.32 ry 22.29 rz -62.41 deg; joints [-4.82, 10.51, 24.35, 0, -29.86, 0] of ABB IRB 5500-27
    - target S4_RBmp2_3 (joint target) at (-863.93, 1912.74, 441.14) mm, rotated rx -168.94 ry 23.92 rz -38.84 deg; joints [20.06, 15.27, 18.02, 0, -28.29, 0] of ABB IRB 5500-27
    - target S4_RBmp3_1 (joint target) at (-871.83, 1930.06, 581.83) mm, rotated rx -168.33 ry 28.01 rz -41.5 deg; joints [20.65, 12.18, 17.28, 0, -24.46, 0] of ABB IRB 5500-27
    - target S4_RBmp3_2 (joint target) at (0.39, 1959.89, 560.27) mm, rotated rx -168.49 ry 26.6 rz -65.21 deg; joints [-4.17, 6.38, 24.38, 0, -25.76, 0] of ABB IRB 5500-27
    - target S4_RBmp3_3 (joint target) at (873.23, 1929.43, 581.83) mm, rotated rx -168.33 ry 28.01 rz -90.16 deg; joints [-28.01, 12.18, 17.28, 0, -24.46, 0] of ABB IRB 5500-27
    - target S4_RBmp4_1 (joint target) at (878.25, 1941.14, 723.32) mm, rotated rx -168.21 ry 32.21 rz -92.9 deg; joints [-27.42, 9.29, 16.35, 0, -20.64, 0] of ABB IRB 5500-27
    - target S4_RBmp4_2 (joint target) at (-0.09, 1952.2, 704.36) mm, rotated rx -168.2 ry 31.08 rz -68.1 deg; joints [-3.52, 2.24, 24.42, 0, -21.66, 0] of ABB IRB 5500-27
    - target S4_RBmp4_3 (joint target) at (-876.96, 1941.72, 723.32) mm, rotated rx -168.21 ry 32.21 rz -44.25 deg; joints [21.23, 9.29, 16.35, 0, -20.64, 0] of ABB IRB 5500-27
    - target S4_Dikki1_1 (joint target) at (910.8, 2059.81, 972.4) mm, rotated rx 177.46 ry 41.17 rz -117.53 deg; joints [-23.24, 9.38, 9.38, 0, 3.24, 0] of ABB IRB 5500-27
    - target S4_Dikki1_2 (joint target) at (99.52, 2054.28, 972.96) mm, rotated rx 177.87 ry 40.72 rz -95.81 deg; joints [-2.18, 0.99, 18.24, 0, 2.76, 0] of ABB IRB 5500-27
    - target S4_Dikki1_3 (joint target) at (-724.17, 2132.59, 972.4) mm, rotated rx 177.46 ry 41.17 rz -74.92 deg; joints [19.37, 9.38, 9.38, 0, 3.24, 0] of ABB IRB 5500-27
    - target S4_Dikki2_1 (joint target) at (-692.33, 2260.68, 1024.72) mm, rotated rx 172.21 ry 42.64 rz -84.13 deg; joints [18.47, 13.4, 3.33, 0, 9.27, 0] of ABB IRB 5500-27
    - target S4_Dikki2_2 (joint target) at (123.49, 2243.77, 1025.17) mm, rotated rx 172.85 ry 42.14 rz -103.42 deg; joints [-1.72, 8.44, 8.88, 0, 8.68, 0] of ABB IRB 5500-27
    - target S4_Dikki2_3 (joint target) at (924.68, 2176, 1024.72) mm, rotated rx 172.21 ry 42.64 rz -124.18 deg; joints [-21.58, 13.4, 3.33, 0, 9.27, 0] of ABB IRB 5500-27
    - target S4_Dikki3_1 (joint target) at (930.8, 2267.3, 1076.08) mm, rotated rx 166.36 ry 43.49 rz -131.4 deg; joints [-20.11, 16.52, -1.85, 0, 15.33, 0] of ABB IRB 5500-27
    - target S4_Dikki3_2 (joint target) at (146.31, 2360.37, 1076.35) mm, rotated rx 167.14 ry 43.08 rz -111.63 deg; joints [-1.34, 12.86, 2.4, 0, 14.73, 0] of ABB IRB 5500-27
    - target S4_Dikki3_3 (joint target) at (-653.35, 2362.24, 1076.08) mm, rotated rx 166.36 ry 43.49 rz -93.62 deg; joints [17.67, 16.52, -1.85, 0, 15.33, 0] of ABB IRB 5500-27
    - target S4_Dikki4_1 (joint target) at (-642.87, 2539.76, 1107.31) mm, rotated rx 159.33 ry 43.89 rz -104 deg; joints [17.08, 23.62, -11.55, 0, 21.93, 0] of ABB IRB 5500-27
    - target S4_Dikki4_2 (joint target) at (168.67, 2460.73, 1121.28) mm, rotated rx 161.01 ry 43.3 rz -120.11 deg; joints [-1.01, 16.83, -3.64, 0, 20.81, 0] of ABB IRB 5500-27
    - target S4_Dikki4_3 (joint target) at (961.27, 2437.14, 1107.31) mm, rotated rx 159.33 ry 43.89 rz -139.73 deg; joints [-18.65, 23.62, -11.55, 0, 21.93, 0] of ABB IRB 5500-27
  - Python program build_cell (listed below)
  - frame Booth_Frame at (0, 1800, 0) mm
    - object Paint_Booth_Floor_12x8m at (0, 0, 0) mm, size 12000 x 8000 x 0 mm
  - frame Rail_Frame at (0, 0, 0) mm
    - object Linear_Track_Bed_7m at (0, 0, 0) mm, size 7000 x 900 x 0 mm
  - frame Car_Frame at (0, 3010, 0) mm
    - object Rotary_Skid_Platform at (0, 0, 0) mm, size 5000 x 2200 x 0 mm
    - object Sedan_Body_4800x1900x1600 at (0, 0, 0) mm, size 4800 x 1900 x 1400 mm
    - object Sedan_Windshields_Glass at (0, 0, 0) mm, size 2860 x 1872.5 x 620 mm
    - object Sedan_Wheels_4x at (0, 0, 0) mm, size 3600 x 1920 x 700 mm
  - program Prog_1_Driver_0deg (74 instructions, listed below)
  - program Prog_2_Front_90deg (31 instructions, listed below)
  - program Prog_3_Passenger_180deg (74 instructions, listed below)
  - program Prog_4_Rear_270deg (28 instructions, listed below)
  - Python program Run_4Stage_Full_Car (listed below)
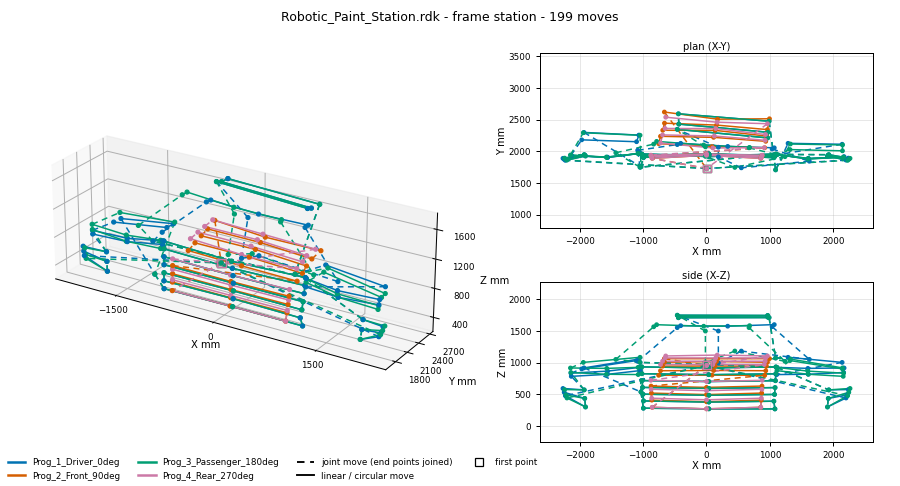
[picture p0: tool path of Robotic_Paint_Station.rdk in frame station, 199 of 199 moves have a stored position in this frame; points joined in program order, loops and branches not executed]

--- Python program build_cell ---
# ==============================================================================
# Final 4-Stage Full-Body Paint Cell (Direct Base Targets + 1880mm MoveL Sweet Spot)
# Candidate: Pavan C S | Assessment: Yuktii AI Labs | Robot: ABB IRB 5500-27
# ==============================================================================
from robolink import *
import math

RDK = Robolink()
RDK.Render(False)

# 1. Connect to ABB Robot and Attached Paint Sprayer Tool
robot = RDK.Item('', ITEM_TYPE_ROBOT)
if not robot.Valid():
    raise Exception("ABB IRB 5500-27 robot not found in station!")

tool = None
for item in robot.Childs():
    if item.Type() == ITEM_TYPE_TOOL:
        tool = item
        break

if tool is None or not tool.Valid():
    raise Exception("Please ensure Generic Paint Sprayer tool is attached!")

# Clean up previous programs, frames, and targets
cleanup_names = [
    'Paint_Full_Cycle', 'Prog_1_Driver_0deg', 'Prog_2_Front_90deg',
    'Prog_3_Passenger_180deg', 'Prog_4_Rear_270deg',
    'Frame_S1_Driver', 'Frame_S2_Front', 'Frame_S3_Passenger', 'Frame_S4_Rear',
    'Car_Frame', 'Booth_Frame', 'Rail_Frame'
]
for name in cleanup_names:
    old = RDK.Item(name)
    if old.Valid():
        old.Delete()

for t in RDK.ItemList(ITEM_TYPE_TARGET):
    t.Delete()

MatClass = robot.Pose().__class__
pi = math.pi

def transl(x, y, z):
    return MatClass([
        [1.0, 0.0, 0.0, float(x)],
        [0.0, 1.0, 0.0, float(y)],
        [0.0, 0.0, 1.0, float(z)],
        [0.0, 0.0, 0.0, 1.0]
    ])

# ==============================================================================
# 2. Exact 25-Point SolveFK Grid (Identical to Working image_f870c6.jpg!)
# ==============================================================================
robot_base = robot.Parent()
robot.setPoseFrame(robot_base)
robot.setPoseTool(tool)
tool_pose = tool.PoseTool()

J2_GRID = [-55.0, -30.0, -5.0, 20.0, 45.0]
J3_GRID = [-42.0, -22.0, -2.0, 18.0, 38.0]

fk_samples = []
for j2_val in J2_GRID:
    for j3_val in J3_GRID:
        j5_val = -(j2_val + j3_val) + 5.0
        tcp = robot.SolveFK([0.0, j2_val, j3_val, 0.0, j5_val, 0.0]) * tool_pose
        fk_samples.append((j2_val, j3_val, tcp[0, 3], tcp[1, 3], tcp[2, 3]))

tcp_j1_test = robot.SolveFK([10.0, -5.0, -2.0, 0.0, 12.0, 0.0]) * tool_pose
tcp_j1_zero = robot.SolveFK([ 0.0, -5.0, -2.0, 0.0, 12.0, 0.0]) * tool_pose
J1_SIGN = 1.0 if (tcp_j1_test[0, 3] < tcp_j1_zero[0, 3]) else -1.0

def solve_exact_from_grid(x_goal, y_goal, z_goal, nozzle_down_deg):
    dpitch = math.radians(nozzle_down_deg - 5.0)
    r_target = math.hypot(x_goal, y_goal) + 160.0 * (1.0 - math.cos(dpitch))
    z_target = z_goal + 210.0 * math.sin(dpitch)

    best_dist = 1e9
    j2_est, j3_est = -5.0, -2.0
    x0_est, y0_est = 174.26, 1880.0
    for (g_j2, g_j3, gx0, gy0, gz0) in fk_samples:
        gr = math.hypot(gx0, gy0)
        d = (gr - r_target)**2 + (gz0 - z_target)**2
        if d < best_dist:
            best_dist = d
            j2_est, j3_est = g_j2, g_j3
            x0_est, y0_est = gx0, gy0

    idx2 = min(len(J2_GRID) - 2, max(0, J2_GRID.index(j2_est)))
    idx3 = min(len(J3_GRID) - 2, max(0, J3_GRID.index(j3_est)))

    def get_cell(i2, i3):
        return fk_samples[i2 * len(J3_GRID) + i3]

    for _ in range(12):
        for k in range(len(J2_GRID) - 1):
            if J2_GRID[k] <= j2_est <= J2_GRID[k+1]:
                idx2 = k
                break
        for k in range(len(J3_GRID) - 1):
            if J3_GRID[k] <= j3_est <= J3_GRID[k+1]:
                idx3 = k
                break

        j2_0, j3_0, x00, y00, z00 = get_cell(idx2, idx3)
        j2_1, _,    x10, y10, z10 = get_cell(idx2 + 1, idx3)
        _,    j3_1, x01, y01, z01 = get_cell(idx2, idx3 + 1)
        _,    _,    x11, y11, z11 = get_cell(idx2 + 1, idx3 + 1)

        r00, r10 = math.hypot(x00, y00), math.hypot(x10, y10)
        r01, r11 = math.hypot(x01, y01), math.hypot(x11, y11)

        u = (j2_est - j2_0) / (j2_1 - j2_0)
        v = (j3_est - j3_0) / (j3_1 - j3_0)

        r_curr = (1-u)*(1-v)*r00 + u*(1-v)*r10 + (1-u)*v*r01 + u*v*r11
        z_curr = (1-u)*(1-v)*z00 + u*(1-v)*z10 + (1-u)*v*z01 + u*v*z11
        x0_est = (1-u)*(1-v)*x00 + u*(1-v)*x10 + (1-u)*v*x01 + u*v*x11
        y0_est = (1-u)*(1-v)*y00 + u*(1-v)*y10 + (1-u)*v*y01 + u*v*y11

        er = r_target - r_curr
        ez = z_target - z_curr
        if abs(er) < 0.3 and abs(ez) < 0.3:
            break

        dr_du = ((1-v)*(r10 - r00) + v*(r11 - r01)) / (j2_1 - j2_0)
        dz_du = ((1-v)*(z10 - z00) + v*(z11 - z01)) / (j2_1 - j2_0)
        dr_dv = ((1-u)*(r01 - r00) + u*(r11 - r10)) / (j3_1 - j3_0)
        dz_dv = ((1-u)*(z01 - z00) + u*(z11 - z10)) / (j3_1 - j3_0)

        det = dr_du * dz_dv - dr_dv * dz_du
        if abs(det) > 1e-3:
            j2_est += 0.8 * (er * dz_dv - dr_dv * ez) / det
            j3_est += 0.8 * (dr_du * ez - er * dz_du) / det

        j2_est = max(-55.0, min(45.0, j2_est))
        j3_est = max(-42.0, min(38.0, j3_est))

    ang_zero = math.degrees(math.atan2(x0_est, y0_est))
    ang_goal = math.degrees(math.atan2(x_goal, y_goal))
    j1 = J1_SIGN * (ang_zero - ang_goal)

    j1 = max(-85.0, min(85.0, j1))
    j5 = max(-65.0, min(65.0, -(j2_est + j3_est) + nozzle_down_deg))
    return [round(j1, 2), round(j2_est, 2), round(j3_est, 2), 0.0, round(j5, 2), 0.0]

# ==============================================================================
# 3. Geometry Setup: Locked Sweet-Spot Distances
# ==============================================================================
DOOR_TCP_Y   = 1880.0
CAR_SIDE_Y   = 3010.0  # 0° & 180° Side Poses: Car side surface at Y=2060, TCP at Y=1880
CAR_END_Y    = 4300.0  # 90° & 270° End Poses: Bumper at 4300-2400 = 1900, Bonnet/Dikki at 1900..2500!

def quad_to_tris(p0, p1, p2, p3):
    return [p0, p1, p2, p0, p2, p3]

def get_car_half_width(z, w_bottom=1900.0, w_top=1520.0, z_cabin_split=920.0):
    if z <= z_cabin_split:
        return w_bottom / 2.0
    factor = (z - z_cabin_split) / (1600.0 - z_cabin_split)
    return (w_bottom / 2.0) * (1.0 - factor) + (w_top / 2.0) * factor

def make_car_along_x(xz_loop, w_bottom, w_top, z_cabin_split=920):
    tris = []
    n = len(xz_loop)
    for i in range(n):
        x1, z1 = xz_loop[i]
        x2, z2 = xz_loop[(i + 1) % n]
        hw1 = get_car_half_width(z1, w_bottom, w_top, z_cabin_split)
        hw2 = get_car_half_width(z2, w_bottom, w_top, z_cabin_split)
        p_f1, p_b1 = [x1, -hw1, z1], [x1, hw1, z1]
        p_f2, p_b2 = [x2, -hw2, z2], [x2, hw2, z2]
        tris.extend(quad_to_tris(p_f1, p_b1, p_b2, p_f2))

    xc, zc = 0.0, 600.0
    hw_c = w_bottom / 2.0
    for i in range(n):
        x1, z1 = xz_loop[i]
        x2, z2 = xz_loop[(i + 1) % n]
        hw1 = get_car_half_width(z1, w_bottom, w_top, z_cabin_split)
        hw2 = get_car_half_width(z2, w_bottom, w_top, z_cabin_split)
        tris.extend([[xc, -hw_c, zc], [x2, -hw2, z2], [x1, -hw1, z1]])
        tris.extend([[xc,  hw_c, zc], [x1,  hw1, z1], [x2,  hw2, z2]])
    return tris

def make_wheel_along_x(x_center, y_in, y_out, z_center, radius=350, segments=24):
    tris = []
    for i in range(segments):
        a1 = 2.0 * pi * i / segments
        a2 = 2.0 * pi * (i + 1) / segments
        x1, z1 = x_center + radius * math.cos(a1), z_center + radius * math.sin(a1)
        x2, z2 = x_center + radius * math.cos(a2), z_center + radius * math.sin(a2)
        tris.extend(quad_to_tris([x1, y_in, z1], [x1, y_out, z1], [x2, y_out, z2], [x2, y_in, z2]))
        tris.extend([[x_center, y_in, z_center], [x2, y_in, z2], [x1, y_in, z1]])
        tris.extend([[x_center, y_out, z_center], [x1, y_out, z1], [x2, y_out, z2]])
    return tris

booth_frame = RDK.AddFrame('Booth_Frame')
booth_frame.setPose(transl(0, 1800, 0))
floor_tris = quad_to_tris([-6000, -4000, 0], [6000, -4000, 0], [6000, 4000, 0], [-6000, 4000, 0])
floor_obj = RDK.AddShape(floor_tris)
floor_obj.setName('Paint_Booth_Floor_12x8m')
floor_obj.setParent(booth_frame)
floor_obj.setColor([0.22, 0.24, 0.27, 0.4])

rail_frame = RDK.AddFrame('Rail_Frame')
rail_frame.setPose(transl(0, 0, 0))
rail_tris = quad_to_tris([-3500, -450, 5], [3500, -450, 5], [3500, 450, 5], [-3500, 450, 5])
rail_obj = RDK.AddShape(rail_tris)
rail_obj.setName('Linear_Track_Bed_7m')
rail_obj.setParent(rail_frame)
rail_obj.setColor([0.75, 0.60, 0.15, 1.0])

car_frame = RDK.AddFrame('Car_Frame')
car_frame.setPose(transl(0, CAR_SIDE_Y, 0))

skid_tris = quad_to_tris([-2500, -1100, 8], [2500, -1100, 8], [2500, 1100, 8], [-2500, 1100, 8])
skid_obj = RDK.AddShape(skid_tris)
skid_obj.setName('Rotary_Skid_Platform')
skid_obj.setParent(car_frame)
skid_obj.setColor([0.35, 0.38, 0.42, 1.0])

sedan_profile = [
    (-2400, 220), (-2400, 520), (-2250, 680), (-1250, 920),
    (-550, 1560), ( 350, 1600), ( 950, 1540), ( 1650, 980),
    ( 2320, 900), ( 2400, 750), ( 2400, 240), ( 1200, 200), (-1200, 200)
]

body_tris = make_car_along_x(sedan_profile, w_bottom=1900.0, w_top=1520.0, z_cabin_split=920.0)
car_body = RDK.AddShape(body_tris)
car_body.setName('Sedan_Body_4800x1900x1600')
car_body.setParent(car_frame)
car_body.setColor([0.18, 0.45, 0.78, 1.0])

glass_tris = []
glass_tris.extend(quad_to_tris([-1230, -760, 930], [-1230, 760, 930], [-560, 680, 1550], [-560, -680, 1550]))
glass_tris.extend(quad_to_tris([ 960, -680, 1530], [ 960, 680, 1530], [ 1630, 760, 990], [ 1630, -760, 990]))

z_win_bot, z_win_top = 980.0, 1450.0
hw_bot = get_car_half_width(z_win_bot) + 3.0
hw_top = get_car_half_width(z_win_top) + 3.0

for side_sign in [-1.0, 1.0]:
    y_wb = side_sign * hw_bot
    y_wt = side_sign * hw_top
    glass_tris.extend(quad_to_tris([-1040.0, y_wb, z_win_bot], [30.0, y_wb, z_win_bot], [30.0, y_wt, z_win_top], [-520.0, y_wt, z_win_top]))
    glass_tris.extend(quad_to_tris([ 210.0, y_wb, z_win_bot], [1380.0, y_wb, z_win_bot], [920.0, y_wt, z_win_top], [ 210.0, y_wt, z_win_top]))

glass_obj = RDK.AddShape(glass_tris)
glass_obj.setName('Sedan_Windshields_Glass')
glass_obj.setParent(car_frame)
glass_obj.setColor([0.12, 0.15, 0.18, 1.0])

wheels_tris = []
for x_axle in [-1450.0, 1450.0]:
    wheels_tris.extend(make_wheel_along_x(x_axle, -960.0, -720.0, 350.0, radius=350.0))
    wheels_tris.extend(make_wheel_along_x(x_axle,  720.0,  960.0, 350.0, radius=350.0))

wheels_obj = RDK.AddShape(wheels_tris)
wheels_obj.setName('Sedan_Wheels_4x')
wheels_obj.setParent(car_frame)
wheels_obj.setColor([0.15, 0.15, 0.15, 1.0])

# ==============================================================================
# 4. Target Generation Parented Directly to robot_base (Zero MoveL Wrist Flip!)
# ==============================================================================
def add_synced_pt(name, x, y, z, nozzle_deg):
    joints = solve_exact_from_grid(x, y, z, nozzle_deg)
    tcp_pose = robot.SolveFK(joints) * tool_pose
    t = RDK.AddTarget(name, robot_base, robot)
    t.setPose(tcp_pose)
    t.setJoints(joints)
    t.setAsJointTarget()
    return t

def add_linear_pass(prog, prefix, x_start, x_end, y_start, y_end, z_start, z_end, nozzle_deg, n_pts=3, use_movej_all=False):
    """
    Point 1 (i == 0) uses MoveJ for row entry; Points 2..N use MoveL for painting!
    Because all targets are in robot_base (just like image_f870c6.jpg), MoveL
    never flips the wrist and never shifts the yellow line away from the arrows!
    """
    for i in range(n_pts):
        f = float(i) / float(n_pts - 1) if n_pts > 1 else 0.0
        x = x_start + f * (x_end - x_start)
        y = y_start + f * (y_end - y_start)
        z = z_start + f * (z_end - z_start)
        pt = add_synced_pt(f"{prefix}_{i+1}", x, y, z, nozzle_deg)
        if use_movej_all or i == 0:
            prog.MoveJ(pt)
        else:
            prog.MoveL(pt)

t_home = add_synced_pt('Target_Home', 0.0, DOOR_TCP_Y - 220.0, 950.0, 5.0)

def build_driver_0_program(prog_name, tag):
    """
    STAGE 1 (0° Driver Side):
    """
    p = RDK.AddProgram(prog_name, robot)
    p.setSpeed(150)
    p.setSpeedJoints(14)
    p.MoveJ(t_home)

    # Zone 1: Front Nose Skirt & Upper Front Fender
    add_linear_pass(p, f'{tag}_Nose1',   -2250, -1860, DOOR_TCP_Y, DOOR_TCP_Y, 320, 320, 5.0, n_pts=2)
    add_linear_pass(p, f'{tag}_Nose2',   -1860, -2250, DOOR_TCP_Y, DOOR_TCP_Y, 450, 450, 5.0, n_pts=2)
    add_linear_pass(p, f'{tag}_Nose3',   -2250, -1860, DOOR_TCP_Y, DOOR_TCP_Y, 580, 580, 5.0, n_pts=2)
    add_linear_pass(p, f'{tag}_Fender1', -2100, -1020, DOOR_TCP_Y, DOOR_TCP_Y, 760, 860, 8.0, n_pts=3)
    add_linear_pass(p, f'{tag}_Fender2', -1020, -2100, DOOR_TCP_Y, DOOR_TCP_Y, 910, 810, 8.0, n_pts=3)
    add_linear_pass(p, f'{tag}_Hood1',   -2000, -1180, DOOR_TCP_Y + 160.0, DOOR_TCP_Y + 160.0, 820, 950, 26.0, n_pts=2)
    add_linear_pass(p, f'{tag}_Hood2',   -1180, -2000, DOOR_TCP_Y + 280.0, DOOR_TCP_Y + 280.0, 970, 840, 30.0, n_pts=2)

    p.MoveJ(add_synced_pt(f'{tag}_Ret_Door', -1000.0, DOOR_TCP_Y - 180.0, 550.0, 5.0))

    # Zone 2: 7-Pass Doors Between Wheels (X = -980 to +1050 mm)
    door_z = [300.0, 405.0, 510.0, 615.0, 720.0, 825.0, 930.0]
    for idx, zv in enumerate(door_z):
        xs, xe = (-980.0, 1050.0) if idx % 2 == 0 else (1050.0, -980.0)
        add_linear_pass(p, f'{tag}_Door{idx+1}', xs, xe, DOOR_TCP_Y, DOOR_TCP_Y, zv, zv, 5.0, n_pts=3)

    p.MoveJ(add_synced_pt(f'{tag}_Ret_Pillar', -1050.0, DOOR_TCP_Y - 180.0, 980.0, 10.0))

    # Zone 3: Greenhouse Pillars
    add_linear_pass(p, f'{tag}_APil', -1120, -540, DOOR_TCP_Y, DOOR_TCP_Y + 145.0,  950, 1490, 22.0, n_pts=2, use_movej_all=True)
    add_linear_pass(p, f'{tag}_Cant',  -520,  920, DOOR_TCP_Y + 165.0, DOOR_TCP_Y + 165.0, 1510, 1510, 28.0, n_pts=3)
    add_linear_pass(p, f'{tag}_CPil',   920, 1520, DOOR_TCP_Y + 145.0, DOOR_TCP_Y, 1490,  980, 22.0, n_pts=2, use_movej_all=True)

    p.MoveJ(add_synced_pt(f'{tag}_Ret_BPil', 500.0, DOOR_TCP_Y - 200.0, 1150.0, 10.0))
    add_linear_pass(p, f'{tag}_BPil',   120,  120, DOOR_TCP_Y, DOOR_TCP_Y + 145.0,  960, 1460, 16.0, n_pts=2, use_movej_all=True)

    # Zone 4: Overhead Left Half-Roof
    add_linear_pass(p, f'{tag}_Roof1', -650,  750, DOOR_TCP_Y + 360.0, DOOR_TCP_Y + 360.0, 1680, 1680, 48.0, n_pts=2)
    add_linear_pass(p, f'{tag}_Roof2',  750, -650, DOOR_TCP_Y + 480.0, DOOR_TCP_Y + 480.0, 1680, 1680, 52.0, n_pts=2)
    add_linear_pass(p, f'{tag}_Roof3', -650,  750, DOOR_TCP_Y + 600.0, DOOR_TCP_Y + 600.0, 1680, 1680, 56.0, n_pts=2)

    p.MoveJ(add_synced_pt(f'{tag}_Ret_Rear', 1050.0, DOOR_TCP_Y - 180.0, 1050.0, 10.0))

    # Zone 5: Left Trunk, Upper Quarter & Rear Skirt
    add_linear_pass(p, f'{tag}_Trnk1', 1150, 2000, DOOR_TCP_Y + 280.0, DOOR_TCP_Y + 280.0, 1000, 930, 28.0, n_pts=2)
    add_linear_pass(p, f'{tag}_Qtr1',  1050, 2100, DOOR_TCP_Y, DOOR_TCP_Y, 800, 820, 8.0, n_pts=3)
    add_linear_pass(p, f'{tag}_Qtr2',  2100, 1050, DOOR_TCP_Y, DOOR_TCP_Y, 890, 910, 8.0, n_pts=3)
    add_linear_pass(p, f'{tag}_RSk1',  1860, 2220, DOOR_TCP_Y, DOOR_TCP_Y, 580, 580, 5.0, n_pts=2)
    add_linear_pass(p, f'{tag}_RSk2',  2220, 1860, DOOR_TCP_Y, DOOR_TCP_Y, 450, 450, 5.0, n_pts=2)
    add_linear_pass(p, f'{tag}_RSk3',  1860, 2220, DOOR_TCP_Y, DOOR_TCP_Y, 320, 320, 5.0, n_pts=2)

    p.MoveJ(t_home)
    return p

def build_passenger_180_program(prog_name, tag):
    """
    STAGE 3 (180° Passenger Side):
    Uses the exact same robot_base parent frame and MoveJ-entry / MoveL-stroke
    pattern as Stage 1!
    """
    p = RDK.AddProgram(prog_name, robot)
    p.setSpeed(150)
    p.setSpeedJoints(14)
    p.MoveJ(t_home)

    # Zone 1: Left Side at 180° (Rear Skirt, Quarter Panel & Right Half-Trunk)
    add_linear_pass(p, f'{tag}_RSk1',  -2220, -1860, DOOR_TCP_Y, DOOR_TCP_Y, 320, 320, 5.0, n_pts=2)
    add_linear_pass(p, f'{tag}_RSk2',  -1860, -2220, DOOR_TCP_Y, DOOR_TCP_Y, 450, 450, 5.0, n_pts=2)
    add_linear_pass(p, f'{tag}_RSk3',  -2220, -1860, DOOR_TCP_Y, DOOR_TCP_Y, 580, 580, 5.0, n_pts=2)
    add_linear_pass(p, f'{tag}_Qtr1',  -2100, -1050, DOOR_TCP_Y, DOOR_TCP_Y, 820, 800, 8.0, n_pts=3)
    add_linear_pass(p, f'{tag}_Qtr2',  -1050, -2100, DOOR_TCP_Y, DOOR_TCP_Y, 910, 890, 8.0, n_pts=3)
    add_linear_pass(p, f'{tag}_Trnk1', -2000, -1150, DOOR_TCP_Y + 280.0, DOOR_TCP_Y + 280.0, 930, 1000, 28.0, n_pts=2)

    p.MoveJ(add_synced_pt(f'{tag}_Ret_Door', -1000.0, DOOR_TCP_Y - 180.0, 550.0, 5.0))

    # Zone 2: 7-Pass Doors Between Wheels (X = -980 to +1050 mm — 100% Wheel-Free!)
    door_z = [300.0, 405.0, 510.0, 615.0, 720.0, 825.0, 930.0]
    for idx, zv in enumerate(door_z):
        xs, xe = (-980.0, 1050.0) if idx % 2 == 0 else (1050.0, -980.0)
        add_linear_pass(p, f'{tag}_Door{idx+1}', xs, xe, DOOR_TCP_Y, DOOR_TCP_Y, zv, zv, 5.0, n_pts=3)

    p.MoveJ(add_synced_pt(f'{tag}_Ret_Pillar', -1050.0, DOOR_TCP_Y - 180.0, 980.0, 10.0))

    # Zone 3: Greenhouse Pillars for 180° (C-Pillar on Left -> Cantrail -> A-Pillar on Right)
    add_linear_pass(p, f'{tag}_CPil', -1480, -900, DOOR_TCP_Y, DOOR_TCP_Y + 145.0,  980, 1490, 22.0, n_pts=2, use_movej_all=True)
    add_linear_pass(p, f'{tag}_Cant',  -880,  540, DOOR_TCP_Y + 165.0, DOOR_TCP_Y + 165.0, 1510, 1510, 28.0, n_pts=3)
    add_linear_pass(p, f'{tag}_APil',   560, 1100, DOOR_TCP_Y + 145.0, DOOR_TCP_Y, 1490,  950, 22.0, n_pts=2, use_movej_all=True)

    p.MoveJ(add_synced_pt(f'{tag}_Ret_BPil', 400.0, DOOR_TCP_Y - 200.0, 1150.0, 10.0))
    add_linear_pass(p, f'{tag}_BPil',   -80,  -80, DOOR_TCP_Y, DOOR_TCP_Y + 145.0,  960, 1460, 16.0, n_pts=2, use_movej_all=True)

    # Zone 4: Overhead Right Half-Roof
    add_linear_pass(p, f'{tag}_Roof1', -650,  750, DOOR_TCP_Y + 360.0, DOOR_TCP_Y + 360.0, 1680, 1680, 48.0, n_pts=2)
    add_linear_pass(p, f'{tag}_Roof2',  750, -650, DOOR_TCP_Y + 480.0, DOOR_TCP_Y + 480.0, 1680, 1680, 52.0, n_pts=2)
    add_linear_pass(p, f'{tag}_Roof3', -650,  750, DOOR_TCP_Y + 600.0, DOOR_TCP_Y + 600.0, 1680, 1680, 56.0, n_pts=2)

    p.MoveJ(add_synced_pt(f'{tag}_Ret_Front', 1050.0, DOOR_TCP_Y - 180.0, 1050.0, 10.0))

    # Zone 5: Right Side at 180° (Right Half-Hood, Front Fender & Front Nose Skirt)
    add_linear_pass(p, f'{tag}_Hood1',  1180, 2000, DOOR_TCP_Y + 280.0, DOOR_TCP_Y + 280.0, 970, 840, 30.0, n_pts=2)
    add_linear_pass(p, f'{tag}_Hood2',  2000, 1180, DOOR_TCP_Y + 160.0, DOOR_TCP_Y + 160.0, 820, 950, 26.0, n_pts=2)
    add_linear_pass(p, f'{tag}_Fend1',  1050, 2100, DOOR_TCP_Y, DOOR_TCP_Y, 860, 760, 8.0, n_pts=3)
    add_linear_pass(p, f'{tag}_Fend2',  2100, 1050, DOOR_TCP_Y, DOOR_TCP_Y, 810, 910, 8.0, n_pts=3)
    add_linear_pass(p, f'{tag}_Nose1',  1860, 2250, DOOR_TCP_Y, DOOR_TCP_Y, 580, 580, 5.0, n_pts=2)
    add_linear_pass(p, f'{tag}_Nose2',  2250, 1860, DOOR_TCP_Y, DOOR_TCP_Y, 450, 450, 5.0, n_pts=2)
    add_linear_pass(p, f'{tag}_Nose3',  1860, 2250, DOOR_TCP_Y, DOOR_TCP_Y, 320, 320, 5.0, n_pts=2)

    p.MoveJ(t_home)
    return p

def build_front_90_program(prog_name, tag):
    """
    STAGE 2 (90° Front Bumper & Bonnet):
    Uses DOOR_TCP_Y = 1880.0 mm for the Bumper and 2020..2480 mm for the Bonnet
    (the exact Y zone that ran without errors in 171157.jpg!), parented to robot_base
    so the yellow path lines sit 100% on the green target arrows!
    """
    p = RDK.AddProgram(prog_name, robot)
    p.setSpeed(150)
    p.setSpeedJoints(14)
    p.MoveJ(t_home)

    # 1. Front Bumper Fascia (4 Full-Width MoveL Sweeps at Y = DOOR_TCP_Y = 1880 mm)
    bmp_z = [300.0, 410.0, 520.0, 630.0]
    for idx, zv in enumerate(bmp_z):
        xs, xe = (-850.0, 850.0) if idx % 2 == 0 else (850.0, -850.0)
        add_linear_pass(p, f'{tag}_Bmp{idx+1}', xs, xe, DOOR_TCP_Y, DOOR_TCP_Y, zv, zv, 5.0, n_pts=3)

    # 2. Front Bonnet / Hood (5 Full-Width MoveL Sweeps from Y = 2000 to Y = 2480 mm)
    bonnet_passes = [
        (DOOR_TCP_Y + 120.0, 740.0, 20.0),
        (DOOR_TCP_Y + 240.0, 800.0, 24.0),
        (DOOR_TCP_Y + 360.0, 860.0, 28.0),
        (DOOR_TCP_Y + 480.0, 920.0, 32.0),
        (DOOR_TCP_Y + 600.0, 970.0, 35.0)
    ]
    for idx, (yv, zv, ang) in enumerate(bonnet_passes):
        xs, xe = (800.0, -800.0) if idx % 2 == 0 else (-800.0, 800.0)
        add_linear_pass(p, f'{tag}_Bonnet{idx+1}', xs, xe, yv, yv, zv, zv, ang, n_pts=3)

    p.MoveJ(t_home)
    return p

def build_rear_270_program(prog_name, tag):
    """
    STAGE 4 (270° Rear Bumper & Back Dikki):
    Uses DOOR_TCP_Y = 1880.0 mm for the Rear Bumper and 2000..2440 mm for the Dikki,
    parented to robot_base so the yellow path lines match the green target arrows!
    """
    p = RDK.AddProgram(prog_name, robot)
    p.setSpeed(150)
    p.setSpeedJoints(14)
    p.MoveJ(t_home)

    # 1. Rear Bumper & Tailgate (4 Full-Width MoveL Sweeps at Y = DOOR_TCP_Y = 1880 mm)
    rear_z = [300.0, 440.0, 580.0, 720.0]
    for idx, zv in enumerate(rear_z):
        xs, xe = (-850.0, 850.0) if idx % 2 == 0 else (850.0, -850.0)
        add_linear_pass(p, f'{tag}_RBmp{idx+1}', xs, xe, DOOR_TCP_Y, DOOR_TCP_Y, zv, zv, 5.0, n_pts=3)

    # 2. Full Back Dikki / Trunk Deck (4 Full-Width MoveL Sweeps from Y = 2000 to Y = 2420 mm)
    dikki_passes = [
        (DOOR_TCP_Y + 120.0,  900.0, 22.0),
        (DOOR_TCP_Y + 260.0,  940.0, 26.0),
        (DOOR_TCP_Y + 400.0,  980.0, 30.0),
        (DOOR_TCP_Y + 540.0, 1020.0, 34.0)
    ]
    for idx, (yv, zv, ang) in enumerate(dikki_passes):
        xs, xe = (780.0, -780.0) if idx % 2 == 0 else (-780.0, 780.0)
        add_linear_pass(p, f'{tag}_Dikki{idx+1}', xs, xe, yv, yv, zv, zv, ang, n_pts=3)

    p.MoveJ(t_home)
    return p

# Build all 4 stage programs:
prog1 = build_driver_0_program('Prog_1_Driver_0deg',          'S1')
prog2 = build_front_90_program('Prog_2_Front_90deg',          'S2')
prog3 = build_passenger_180_program('Prog_3_Passenger_180deg', 'S3')
prog4 = build_rear_270_program('Prog_4_Rear_270deg',          'S4')

# Hide S2, S3, S4 targets initially so only Pose 1 targets are shown
for t in RDK.ItemList(ITEM_TYPE_TARGET):
    tname = t.Name()
    t.setVisible(tname.startswith('S1_') or tname == 'Target_Home')

robot.setJoints(t_home.Joints())
RDK.Render(True)
print("SUCCESS: All 4 Poses Built Directly in robot_base (Zero Shift + Zero Popups)!")

--- program Prog_1_Driver_0deg (robot ABB IRB 5500-27) ---
  Set speed (150.0 mm/s)
  Set speed (14.0 deg/s)
  MoveJ (Target_Home)
  MoveJ (S1_Nose1_1)
  MoveL (S1_Nose1_2)
  MoveJ (S1_Nose2_1)
  MoveL (S1_Nose2_2)
  MoveJ (S1_Nose3_1)
  MoveL (S1_Nose3_2)
  MoveJ (S1_Fender1_1)
  MoveL (S1_Fender1_2)
  MoveL (S1_Fender1_3)
  MoveJ (S1_Fender2_1)
  MoveL (S1_Fender2_2)
  MoveL (S1_Fender2_3)
  MoveJ (S1_Hood1_1)
  MoveL (S1_Hood1_2)
  MoveJ (S1_Hood2_1)
  MoveL (S1_Hood2_2)
  MoveJ (S1_Ret_Door)
  MoveJ (S1_Door1_1)
  MoveL (S1_Door1_2)
  MoveL (S1_Door1_3)
  MoveJ (S1_Door2_1)
  MoveL (S1_Door2_2)
  MoveL (S1_Door2_3)
  MoveJ (S1_Door3_1)
  MoveL (S1_Door3_2)
  MoveL (S1_Door3_3)
  MoveJ (S1_Door4_1)
  MoveL (S1_Door4_2)
  MoveL (S1_Door4_3)
  MoveJ (S1_Door5_1)
  MoveL (S1_Door5_2)
  MoveL (S1_Door5_3)
  MoveJ (S1_Door6_1)
  MoveL (S1_Door6_2)
  MoveL (S1_Door6_3)
  MoveJ (S1_Door7_1)
  MoveL (S1_Door7_2)
  MoveL (S1_Door7_3)
  MoveJ (S1_Ret_Pillar)
  MoveJ (S1_APil_1)
  MoveJ (S1_APil_2)
  MoveJ (S1_Cant_1)
  MoveL (S1_Cant_2)
  MoveL (S1_Cant_3)
  MoveJ (S1_CPil_1)
  MoveJ (S1_CPil_2)
  MoveJ (S1_Ret_BPil)
  MoveJ (S1_BPil_1)
  MoveJ (S1_BPil_2)
  MoveJ (S1_Roof1_1)
  MoveL (S1_Roof1_2)
  MoveJ (S1_Roof2_1)
  MoveL (S1_Roof2_2)
  MoveJ (S1_Roof3_1)
  MoveL (S1_Roof3_2)
  MoveJ (S1_Ret_Rear)
  MoveJ (S1_Trnk1_1)
  MoveL (S1_Trnk1_2)
  MoveJ (S1_Qtr1_1)
  MoveL (S1_Qtr1_2)
  MoveL (S1_Qtr1_3)
  MoveJ (S1_Qtr2_1)
  MoveL (S1_Qtr2_2)
  MoveL (S1_Qtr2_3)
  MoveJ (S1_RSk1_1)
  MoveL (S1_RSk1_2)
  MoveJ (S1_RSk2_1)
  MoveL (S1_RSk2_2)
  MoveJ (S1_RSk3_1)
  MoveL (S1_RSk3_2)
  MoveJ (Target_Home)

--- program Prog_2_Front_90deg (robot ABB IRB 5500-27) ---
  Set speed (150.0 mm/s)
  Set speed (14.0 deg/s)
  MoveJ (Target_Home)
  MoveJ (S2_Bmp1_1)
  MoveL (S2_Bmp1_2)
  MoveL (S2_Bmp1_3)
  MoveJ (S2_Bmp2_1)
  MoveL (S2_Bmp2_2)
  MoveL (S2_Bmp2_3)
  MoveJ (S2_Bmp3_1)
  MoveL (S2_Bmp3_2)
  MoveL (S2_Bmp3_3)
  MoveJ (S2_Bmp4_1)
  MoveL (S2_Bmp4_2)
  MoveL (S2_Bmp4_3)
  MoveJ (S2_Bonnet1_1)
  MoveL (S2_Bonnet1_2)
  MoveL (S2_Bonnet1_3)
  MoveJ (S2_Bonnet2_1)
  MoveL (S2_Bonnet2_2)
  MoveL (S2_Bonnet2_3)
  MoveJ (S2_Bonnet3_1)
  MoveL (S2_Bonnet3_2)
  MoveL (S2_Bonnet3_3)
  MoveJ (S2_Bonnet4_1)
  MoveL (S2_Bonnet4_2)
  MoveL (S2_Bonnet4_3)
  MoveJ (S2_Bonnet5_1)
  MoveL (S2_Bonnet5_2)
  MoveL (S2_Bonnet5_3)
  MoveJ (Target_Home)

--- program Prog_3_Passenger_180deg (robot ABB IRB 5500-27) ---
  Set speed (150.0 mm/s)
  Set speed (14.0 deg/s)
  MoveJ (Target_Home)
  MoveJ (S3_RSk1_1)
  MoveL (S3_RSk1_2)
  MoveJ (S3_RSk2_1)
  MoveL (S3_RSk2_2)
  MoveJ (S3_RSk3_1)
  MoveL (S3_RSk3_2)
  MoveJ (S3_Qtr1_1)
  MoveL (S3_Qtr1_2)
  MoveL (S3_Qtr1_3)
  MoveJ (S3_Qtr2_1)
  MoveL (S3_Qtr2_2)
  MoveL (S3_Qtr2_3)
  MoveJ (S3_Trnk1_1)
  MoveL (S3_Trnk1_2)
  MoveJ (S3_Ret_Door)
  MoveJ (S3_Door1_1)
  MoveL (S3_Door1_2)
  MoveL (S3_Door1_3)
  MoveJ (S3_Door2_1)
  MoveL (S3_Door2_2)
  MoveL (S3_Door2_3)
  MoveJ (S3_Door3_1)
  MoveL (S3_Door3_2)
  MoveL (S3_Door3_3)
  MoveJ (S3_Door4_1)
  MoveL (S3_Door4_2)
  MoveL (S3_Door4_3)
  MoveJ (S3_Door5_1)
  MoveL (S3_Door5_2)
  MoveL (S3_Door5_3)
  MoveJ (S3_Door6_1)
  MoveL (S3_Door6_2)
  MoveL (S3_Door6_3)
  MoveJ (S3_Door7_1)
  MoveL (S3_Door7_2)
  MoveL (S3_Door7_3)
  MoveJ (S3_Ret_Pillar)
  MoveJ (S3_CPil_1)
  MoveJ (S3_CPil_2)
  MoveJ (S3_Cant_1)
  MoveL (S3_Cant_2)
  MoveL (S3_Cant_3)
  MoveJ (S3_APil_1)
  MoveJ (S3_APil_2)
  MoveJ (S3_Ret_BPil)
  MoveJ (S3_BPil_1)
  MoveJ (S3_BPil_2)
  MoveJ (S3_Roof1_1)
  MoveL (S3_Roof1_2)
  MoveJ (S3_Roof2_1)
  MoveL (S3_Roof2_2)
  MoveJ (S3_Roof3_1)
  MoveL (S3_Roof3_2)
  MoveJ (S3_Ret_Front)
  MoveJ (S3_Hood1_1)
  MoveL (S3_Hood1_2)
  MoveJ (S3_Hood2_1)
  MoveL (S3_Hood2_2)
  MoveJ (S3_Fend1_1)
  MoveL (S3_Fend1_2)
  MoveL (S3_Fend1_3)
  MoveJ (S3_Fend2_1)
  MoveL (S3_Fend2_2)
  MoveL (S3_Fend2_3)
  MoveJ (S3_Nose1_1)
  MoveL (S3_Nose1_2)
  MoveJ (S3_Nose2_1)
  MoveL (S3_Nose2_2)
  MoveJ (S3_Nose3_1)
  MoveL (S3_Nose3_2)
  MoveJ (Target_Home)

--- program Prog_4_Rear_270deg (robot ABB IRB 5500-27) ---
  Set speed (150.0 mm/s)
  Set speed (14.0 deg/s)
  MoveJ (Target_Home)
  MoveJ (S4_RBmp1_1)
  MoveL (S4_RBmp1_2)
  MoveL (S4_RBmp1_3)
  MoveJ (S4_RBmp2_1)
  MoveL (S4_RBmp2_2)
  MoveL (S4_RBmp2_3)
  MoveJ (S4_RBmp3_1)
  MoveL (S4_RBmp3_2)
  MoveL (S4_RBmp3_3)
  MoveJ (S4_RBmp4_1)
  MoveL (S4_RBmp4_2)
  MoveL (S4_RBmp4_3)
  MoveJ (S4_Dikki1_1)
  MoveL (S4_Dikki1_2)
  MoveL (S4_Dikki1_3)
  MoveJ (S4_Dikki2_1)
  MoveL (S4_Dikki2_2)
  MoveL (S4_Dikki2_3)
  MoveJ (S4_Dikki3_1)
  MoveL (S4_Dikki3_2)
  MoveL (S4_Dikki3_3)
  MoveJ (S4_Dikki4_1)
  MoveL (S4_Dikki4_2)
  MoveL (S4_Dikki4_3)
  MoveJ (Target_Home)

--- Python program Run_4Stage_Full_Car ---
from robolink import *
import math
import time
import tkinter as tk
from tkinter import simpledialog

RDK = Robolink()
car_frame = RDK.Item('Car_Frame', ITEM_TYPE_FRAME)
MatClass = car_frame.Pose().__class__

CAR_SIDE_Y = 3010.0  # Locked for 0° and 180°
CAR_END_Y  = 4300.0  # Locked for 90° and 270° (Places Bumper at Y=1900, TCP at 1880!)

def show_only_prefix(prefix):
    """Shows ONLY targets starting with 'S1_', 'S2_', 'S3_', or 'S4_' so screen is clean!"""
    RDK.Render(False)
    for t in RDK.ItemList(ITEM_TYPE_TARGET):
        tname = t.Name()
        t.setVisible(tname.startswith(prefix) or tname == 'Target_Home')
    RDK.Render(True)

def set_car_pose(deg, y_pos):
    ang = math.radians(deg)
    ca, sa = float(math.cos(ang)), float(math.sin(ang))
    car_frame.setPose(MatClass([
        [ca, -sa, 0.0, 0.0],
        [sa,  ca, 0.0, float(y_pos)],
        [0.0, 0.0, 1.0, 0.0],
        [0.0, 0.0, 0.0, 1.0]
    ]))

def animate_turntable(start_deg, end_deg, y_start, y_end):
    for step in range(25):
        f = step / 24.0
        set_car_pose(start_deg + f * (end_deg - start_deg), y_start + f * (y_end - y_start))
        time.sleep(0.03)

def run_stage_blocking(prog_name):
    p = RDK.Item(prog_name, ITEM_TYPE_PROGRAM)
    if p.Valid():
        p.RunProgram()
        while p.Busy():
            time.sleep(0.1)

root = tk.Tk()
root.withdraw()
root.attributes("-topmost", True)
choice = simpledialog.askstring(
    "Select Pose to Run",
    "Enter Pose Number (0, 1, 2, 3, or 4):\n\n"
    "0 = Run ALL 4 Poses Together (Full 360° Car)\n"
    "1 = Pose 1 ONLY (0° Driver Side)\n"
    "2 = Pose 2 ONLY (90° Front Bumper & Bonnet)\n"
    "3 = Pose 3 ONLY (180° Passenger Side)\n"
    "4 = Pose 4 ONLY (270° Rear Bumper & Back Dikki)",
    initialvalue="0",
    parent=root
)
root.destroy()

if choice is not None:
    mode = str(choice).strip()

    if mode == "1":
        show_only_prefix('S1_')
        set_car_pose(0.0, CAR_SIDE_Y)
        run_stage_blocking('Prog_1_Driver_0deg')

    elif mode == "2":
        show_only_prefix('S2_')
        set_car_pose(90.0, CAR_END_Y)
        run_stage_blocking('Prog_2_Front_90deg')

    elif mode == "3":
        show_only_prefix('S3_')
        set_car_pose(180.0, CAR_SIDE_Y)
        run_stage_blocking('Prog_3_Passenger_180deg')

    elif mode == "4":
        show_only_prefix('S4_')
        set_car_pose(270.0, CAR_END_Y)
        run_stage_blocking('Prog_4_Rear_270deg')

    elif mode == "0":
        show_only_prefix('S1_')
        set_car_pose(0.0, CAR_SIDE_Y)
        run_stage_blocking('Prog_1_Driver_0deg')

        animate_turntable(0.0, 90.0, CAR_SIDE_Y, CAR_END_Y)
        show_only_prefix('S2_')
        run_stage_blocking('Prog_2_Front_90deg')

        animate_turntable(90.0, 180.0, CAR_END_Y, CAR_SIDE_Y)
        show_only_prefix('S3_')
        run_stage_blocking('Prog_3_Passenger_180deg')

        animate_turntable(180.0, 270.0, CAR_SIDE_Y, CAR_END_Y)
        show_only_prefix('S4_')
        run_stage_blocking('Prog_4_Rear_270deg')

        animate_turntable(270.0, 360.0, CAR_END_Y, CAR_SIDE_Y)
        show_only_prefix('S1_')
